PROGRAM PersistentCaller
VAR
	persistanceHandler : FB_PersistentHandler;
	enable	: BOOL := TRUE;
	reinit	: BOOL := FALSE;
END_VAR


persistanceHandler(bEnable := enable,
				   bReinit := reinit);

END_PROGRAM

(* stored: Version 1.1.0.1
   POU PersistentCaller: Id {1d6c7289-79d4-45ba-a765-47310686d7f4}, SpecialFunc None *)
